FUNCTION_BLOCK fbRoomLiving IMPLEMENTS iRoom
VAR
	
//  ----------- RELAYS -----------
	ShutterR1OpenRelay : fbMonostableRelay;
	ShutterR1CloseRelay : fbMonostableRelay;
	LightH1Relay : fbBistableSingleCoilRelay;
	
//  ----------- SWITCHES -----------
	ShutterR1OpenSwitch : fbMonoSwitch;
	ShutterR1CloseSwitch : fbMonoSwitch;
	LightH1Switch : fbMonoSwitch;
	
//  ----------- SWITCH CONTROLLERS -----------	
	ShutterR1OpenSwitchCtrl : fbSwitchCtrl;	
	ShutterR1CloseSwitchCtrl : fbSwitchCtrl;	
	LightH1SwitchCtrl : fbSwitchCtrl;											

	
//  ----------- SHUTTER CONTROLLERS -----------	
	ShutterR1Ctrl : fbShutterCtrl;
	
//  ----------- LIGHT CONTROLLERS -----------	
	LightH1Ctrl : fbLightCtrl;	
	
	
//  ----------- SHUTTER CMD SOURCES -----------
	ShutterR1CmdEvent : stShutterCmdEvent;
	ShutterR1CmdSwitch : fbShutterCmdSourceSwitch;
	ShutterR1CmdHa : fbShutterCmdSourceHa;
	
//  ----------- SHUTTER CMD SOURCES -----------
	LightH1CmdEvent : stLightCmdEvent;
END_VAR


//  ----------- RUN SWITCHES -----------	
ShutterR1OpenSwitch();
ShutterR1CloseSwitch();
LightH1Switch();

//  ----------- RUN SWITCH CONTROLLERS -----------
ShutterR1OpenSwitchCtrl(Switch := ShutterR1OpenSwitch,
						Config := gvlSwitches.GeneralSwitchConfig);
ShutterR1CloseSwitchCtrl(Switch := ShutterR1CloseSwitch,
						Config := gvlSwitches.GeneralSwitchConfig);


//  ----------- RUN SHUTTER CMD SOURCES -----------
ShutterR1CmdSwitch( OpenSwitchState := ShutterR1OpenSwitchCtrl.State,
						CloseSwitchState := ShutterR1CloseSwitchCtrl.State,
						ShutterStateType := ShutterR1Ctrl.CurrentState.StateType,
						ShutterConfig := gvlShutters.ShutterR1Config);
ShutterR1CmdSwitch.Process(CmdEvent := ShutterR1CmdEvent);

ShutterR1CmdHa( HaCmdEvent := gvlHA.Shutter1CmdEvent) ;
ShutterR1CmdHa.Process(CmdEvent := ShutterR1CmdEvent);



//  ----------- RUN SHUTTER CONTROLLERS -----------
ShutterR1Ctrl(ShutterOpenRelay := ShutterR1OpenRelay,
			ShutterCloseRelay := ShutterR1CloseRelay,
			ShutterConfig := gvlShutters.ShutterR1Config,
			CmdEvent := ShutterR1CmdEvent);

//  ----------- RUN LIGHT CONTROLLERS -----------
LightH1Ctrl( LightRelay :=LightH1Relay,
				Config := gvlLights.LightH1Config,
				Smoothing := TRUE,
				State :=,
				Brightness :=,
				CmdEvent := );

METHOD LightsOff
// Light1Ctrl.TurnOff();
// Light2Ctrl.TurnOff();
// Light3Ctrl.TurnOff();
END_METHOD

METHOD LightsOn
// Light1Ctrl.TurnOn();
// Light2Ctrl.TurnOn();
// Light3Ctrl.TurnOn();
END_METHOD

METHOD ShuttersClose
END_METHOD

METHOD ShuttersOpen
END_METHOD

END_FUNCTION_BLOCK

(* stored: Version 1.1.0.1
   POU fbRoomLiving: Id {74a16cd5-868a-413e-b1b4-1075b610be2f}, SpecialFunc None
   Method LightsOff: Id {262cd78d-a037-4ac4-890b-0001e3f12830}
   Method LightsOn: Id {ff3dfedc-8e50-4daa-a0a5-a2f01180a960}
   Method ShuttersClose: Id {fb9fcdd0-daee-4038-9b3b-8a88f7bea9a5}
   Method ShuttersOpen: Id {d21a0eb5-595a-4dea-8b06-37dc33bd6a36} *)
